Fanuc KAREL source: KA00003.KL

PROGRAM KA00003
%NOLOCKGROUP
VAR
  SRC: INTEGER
  DST: BOOLEAN
BEGIN
  SRC = 2
  DST = SRC
END KA00003
